// TIA Portal V21 export
// export: Created 2000-01-01T00:00:00.0000000Z, ExportSetting None
FUNCTION "MCP_B6_LadFc" : Void   // FC9602, LAD
TITLE = 条件与定时
{ S7_Optimized_Access := 'TRUE' }
// stored: SetENOAutomatically false
BEGIN

REGION Network 1
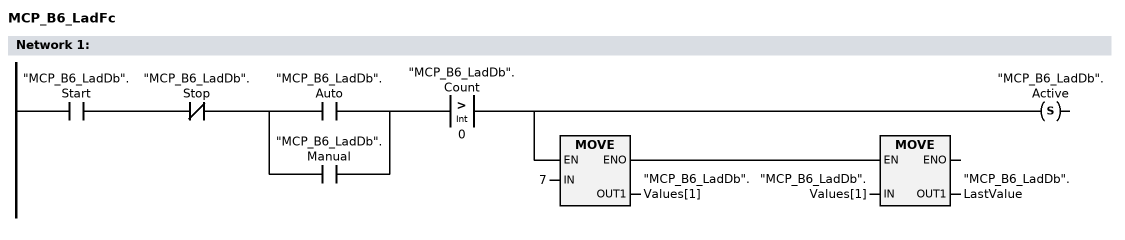
   RUNG wire#powerrail
      Contact( "MCP_B6_LadDb".Start )
      I_Contact( "MCP_B6_LadDb".Stop )
      wire#w1
      Contact( "MCP_B6_LadDb".Auto )
      wire#w2
      { S7_Templates := "SrcType := Int" } GT_Contact(in1 := "MCP_B6_LadDb".Count, in2 := 0)
      wire#w3
      S_Coil( "MCP_B6_LadDb".Active )
   END_RUNG
   RUNG wire#w1
      Contact( "MCP_B6_LadDb".Manual )
   END_RUNG wire#w2
   RUNG wire#w3
      { S7_GenerateENO := "TRUE" } Move(in := 7, out1 => "MCP_B6_LadDb".Values[1])
      Move(in := "MCP_B6_LadDb".Values[1], out1 => "MCP_B6_LadDb".LastValue)
   END_RUNG
   // the same network as SCL:
   // ENO of a box is taken as its EN; it also drops when the box reports an error
   IF "MCP_B6_LadDb".Start AND NOT "MCP_B6_LadDb".Stop AND ("MCP_B6_LadDb".Auto OR "MCP_B6_LadDb".Manual) AND ("MCP_B6_LadDb".Count > 0) THEN
       "MCP_B6_LadDb".Active := TRUE;
       "MCP_B6_LadDb".Values[1] := 7;
       "MCP_B6_LadDb".LastValue := "MCP_B6_LadDb".Values[1];
   END_IF;
END_REGION
END_FUNCTION
